// Tests for HalfBROT.F_FocusTargetFollowsActual (HalfBROT 0.7.2): the focus target follows the actual position after a hand move.
FUNCTION_BLOCK F_FocusTargetFollowsActual_Tests EXTENDS TcUnit.FB_TestSuite
VAR
END_VAR

Manual_Calibrated_Follows();
Automatic_Idle_Does_Not_Follow();
Automatic_Jogging_Follows();
Not_Calibrated_Never();
Homing_Never();

// Manual or off mode: the pendant moves the focus, the target follows it.
METHOD PRIVATE Manual_Calibrated_Follows
VAR
END_VAR
TEST('Manual_Calibrated_Follows');
AssertTrue(Condition := HalfBROT.F_FocusTargetFollowsActual(bAutomatic := FALSE, bManualUnlock := FALSE, bJogging := FALSE, bCalibrated := TRUE, bHoming := FALSE), Message := 'manual or off, calibrated');
TEST_FINISHED();
END_METHOD

// Automatic positioning owns the target.
METHOD PRIVATE Automatic_Idle_Does_Not_Follow
VAR
END_VAR
TEST('Automatic_Idle_Does_Not_Follow');
AssertFalse(Condition := HalfBROT.F_FocusTargetFollowsActual(bAutomatic := TRUE, bManualUnlock := FALSE, bJogging := FALSE, bCalibrated := TRUE, bHoming := FALSE), Message := 'automatic, idle');
TEST_FINISHED();
END_METHOD

// A pendant jog in automatic mode (the pendant is not mode gated) and a manual unlock also move the focus by hand.
METHOD PRIVATE Automatic_Jogging_Follows
VAR
END_VAR
TEST('Automatic_Jogging_Follows');
AssertTrue(Condition := HalfBROT.F_FocusTargetFollowsActual(bAutomatic := TRUE, bManualUnlock := FALSE, bJogging := TRUE, bCalibrated := TRUE, bHoming := FALSE), Message := 'automatic, jogging');
AssertTrue(Condition := HalfBROT.F_FocusTargetFollowsActual(bAutomatic := TRUE, bManualUnlock := TRUE, bJogging := FALSE, bCalibrated := TRUE, bHoming := FALSE), Message := 'automatic, manual unlock');
TEST_FINISHED();
END_METHOD

// An uncalibrated focus has no actual position to follow, in any mode.
METHOD PRIVATE Not_Calibrated_Never
VAR
END_VAR
TEST('Not_Calibrated_Never');
AssertFalse(Condition := HalfBROT.F_FocusTargetFollowsActual(bAutomatic := FALSE, bManualUnlock := FALSE, bJogging := FALSE, bCalibrated := FALSE, bHoming := FALSE), Message := 'not calibrated, a=FALSE u=FALSE j=FALSE');
AssertFalse(Condition := HalfBROT.F_FocusTargetFollowsActual(bAutomatic := FALSE, bManualUnlock := FALSE, bJogging := TRUE, bCalibrated := FALSE, bHoming := FALSE), Message := 'not calibrated, a=FALSE u=FALSE j=TRUE');
AssertFalse(Condition := HalfBROT.F_FocusTargetFollowsActual(bAutomatic := FALSE, bManualUnlock := TRUE, bJogging := FALSE, bCalibrated := FALSE, bHoming := FALSE), Message := 'not calibrated, a=FALSE u=TRUE j=FALSE');
AssertFalse(Condition := HalfBROT.F_FocusTargetFollowsActual(bAutomatic := FALSE, bManualUnlock := TRUE, bJogging := TRUE, bCalibrated := FALSE, bHoming := FALSE), Message := 'not calibrated, a=FALSE u=TRUE j=TRUE');
AssertFalse(Condition := HalfBROT.F_FocusTargetFollowsActual(bAutomatic := TRUE, bManualUnlock := FALSE, bJogging := FALSE, bCalibrated := FALSE, bHoming := FALSE), Message := 'not calibrated, a=TRUE u=FALSE j=FALSE');
AssertFalse(Condition := HalfBROT.F_FocusTargetFollowsActual(bAutomatic := TRUE, bManualUnlock := FALSE, bJogging := TRUE, bCalibrated := FALSE, bHoming := FALSE), Message := 'not calibrated, a=TRUE u=FALSE j=TRUE');
AssertFalse(Condition := HalfBROT.F_FocusTargetFollowsActual(bAutomatic := TRUE, bManualUnlock := TRUE, bJogging := FALSE, bCalibrated := FALSE, bHoming := FALSE), Message := 'not calibrated, a=TRUE u=TRUE j=FALSE');
AssertFalse(Condition := HalfBROT.F_FocusTargetFollowsActual(bAutomatic := TRUE, bManualUnlock := TRUE, bJogging := TRUE, bCalibrated := FALSE, bHoming := FALSE), Message := 'not calibrated, a=TRUE u=TRUE j=TRUE');
TEST_FINISHED();
END_METHOD

// The homing owns fPosition, in any mode.
METHOD PRIVATE Homing_Never
VAR
END_VAR
TEST('Homing_Never');
AssertFalse(Condition := HalfBROT.F_FocusTargetFollowsActual(bAutomatic := FALSE, bManualUnlock := FALSE, bJogging := FALSE, bCalibrated := TRUE, bHoming := TRUE), Message := 'homing, a=FALSE u=FALSE j=FALSE');
AssertFalse(Condition := HalfBROT.F_FocusTargetFollowsActual(bAutomatic := FALSE, bManualUnlock := FALSE, bJogging := TRUE, bCalibrated := TRUE, bHoming := TRUE), Message := 'homing, a=FALSE u=FALSE j=TRUE');
AssertFalse(Condition := HalfBROT.F_FocusTargetFollowsActual(bAutomatic := FALSE, bManualUnlock := TRUE, bJogging := FALSE, bCalibrated := TRUE, bHoming := TRUE), Message := 'homing, a=FALSE u=TRUE j=FALSE');
AssertFalse(Condition := HalfBROT.F_FocusTargetFollowsActual(bAutomatic := FALSE, bManualUnlock := TRUE, bJogging := TRUE, bCalibrated := TRUE, bHoming := TRUE), Message := 'homing, a=FALSE u=TRUE j=TRUE');
AssertFalse(Condition := HalfBROT.F_FocusTargetFollowsActual(bAutomatic := TRUE, bManualUnlock := FALSE, bJogging := FALSE, bCalibrated := TRUE, bHoming := TRUE), Message := 'homing, a=TRUE u=FALSE j=FALSE');
AssertFalse(Condition := HalfBROT.F_FocusTargetFollowsActual(bAutomatic := TRUE, bManualUnlock := FALSE, bJogging := TRUE, bCalibrated := TRUE, bHoming := TRUE), Message := 'homing, a=TRUE u=FALSE j=TRUE');
AssertFalse(Condition := HalfBROT.F_FocusTargetFollowsActual(bAutomatic := TRUE, bManualUnlock := TRUE, bJogging := FALSE, bCalibrated := TRUE, bHoming := TRUE), Message := 'homing, a=TRUE u=TRUE j=FALSE');
AssertFalse(Condition := HalfBROT.F_FocusTargetFollowsActual(bAutomatic := TRUE, bManualUnlock := TRUE, bJogging := TRUE, bCalibrated := TRUE, bHoming := TRUE), Message := 'homing, a=TRUE u=TRUE j=TRUE');
TEST_FINISHED();
END_METHOD

END_FUNCTION_BLOCK

(* stored: Version 1.1.0.1, ProductVersion 3.1.4024.15
   POU F_FocusTargetFollowsActual_Tests: Id {124fa07e-a7a8-4d27-ae7a-5ed8dbb24aca}, SpecialFunc None
   Method Manual_Calibrated_Follows: Id {16f0bdbc-9e3f-41cd-97fa-0a533b59b994}
   Method Automatic_Idle_Does_Not_Follow: Id {522384bc-f9d8-4e55-af6f-b3f6066da3a8}
   Method Automatic_Jogging_Follows: Id {c644cadb-7db0-4aed-a77d-10a74a0e88e4}
   Method Not_Calibrated_Never: Id {e200a10a-4dcd-4217-ae20-0a7ab579c3e2}
   Method Homing_Never: Id {fd66d9ef-7416-4653-882c-9612fec1989b} *)
